(* IEC 61131-3 sources: avi-aoi-management/scripts/ai-eval/ngau-nhien/kho/st-tt1-bo-phieu-2oo3/mau/src, 1 file *)

(* ---- BoPhieu2oo3.st ---- *)
FUNCTION_BLOCK BoPhieu2oo3
VAR_INPUT
    A : BOOL;
    B : BOOL;
    C : BOOL;
    RESET : BOOL;
END_VAR
VAR_OUTPUT
    Q : BOOL;
    LECH : BOOL;
    KENH_LECH : INT;
    DEM_LECH : DINT;
END_VAR
VAR
    lechCu : BOOL;
    soTrue : INT;
END_VAR
    soTrue := BOOL_TO_INT(A) + BOOL_TO_INT(B) + BOOL_TO_INT(C);
    Q := soTrue >= 2;
    LECH := (soTrue = 1) OR (soTrue = 2);
    IF NOT LECH THEN
        KENH_LECH := 0;
    ELSIF soTrue = 1 THEN
        (* kênh lệch là kênh TRUE duy nhất *)
        IF A THEN KENH_LECH := 1; ELSIF B THEN KENH_LECH := 2; ELSE KENH_LECH := 3; END_IF
    ELSE
        (* kênh lệch là kênh FALSE duy nhất *)
        IF NOT A THEN KENH_LECH := 1; ELSIF NOT B THEN KENH_LECH := 2; ELSE KENH_LECH := 3; END_IF
    END_IF
    IF RESET THEN
        DEM_LECH := 0;
    ELSIF LECH AND NOT lechCu THEN
        DEM_LECH := DEM_LECH + 1;
    END_IF
    lechCu := LECH;
END_FUNCTION_BLOCK
